(* IEC 61131-3 sources: codesys-framework/txt/application/WeVe Core (library)/70 Logger, 1 file *)

(* ---- GVL_Logger.gvl.st ---- *)
{attribute 'qualified_only'}
VAR_GLOBAL CONSTANT
	cMaxMessageLength 	: UINT := 255;		// max lengte van een gelogde boodschap
END_VAR
